// TIA Portal V20 export
// export: Created 2026-10-20T12:44:55.4293311Z, ExportSetting WithDefaults, DisplayName Totally Integrated Automation Portal, DisplayVersion V20 Update 6, DisplayName TIA Portal Openness, DisplayVersion V20 Update 6, DisplayName TIA Portal Version Control Interface, DisplayVersion V20 Update 6, DisplayName SINAMICS Startdrive Advanced, DisplayVersion V20 SP1, DisplayName SINAMICS Startdrive G130, G150, S120, S150, SINAMICS MV, G220, S200, S210, DisplayVersion V20 SP1, DisplayName SINAMICS Startdrive G110M, G120, G120C, G120D, G120P, G115D, DisplayVersion V20 SP1, DisplayName STEP 7 Professional, DisplayVersion V20 Update 6, DisplayName STEP 7 Safety, DisplayVersion V20 Update 2, DisplayName WinCC Basic/Comfort/Advanced, DisplayVersion V20 Update 6, DisplayName WinCC Unified, DisplayVersion V20 Update 6
FUNCTION "CNV_Selector_1" : Void   // FC60, SCL
{ S7_Optimized_Access := 'TRUE' }
VERSION : 0.1
// stored: AutoNumber true, IsIECCheckEnabled false, SetENOAutomatically false, UDAEnableTagReadback false
   VAR_INPUT
      Sys_No : UInt;
      Zone : UInt;
      CNV1_2_Selected : UInt;
   END_VAR
   VAR_OUTPUT
      ID : DInt;
      "ID(1)" : DInt;
   END_VAR
BEGIN
   //CNV SCREEN SELECTION
   CASE #Sys_No OF
       0:
           #ID := 0;
           #"ID(1)" := 0;

       1://SYSTEM 1
           #ID := "Settings_DB".ECnv_Sys[1].ID; // EXTRACTOR CONVEYOR
           CASE #Zone OF
               11: //LEVEL 1
                   IF #CNV1_2_Selected = 1 THEN
                       #"ID(1)" := "Settings_DB".LCnv_Sys[1].Cnv_Level[1].Cnv1.ID; //CNV 1
                   ELSIF #CNV1_2_Selected = 2 THEN
                       #"ID(1)" := "Settings_DB".LCnv_Sys[1].Cnv_Level[1].Cnv2.ID; //CNV 2
                   END_IF;
               12: //LEVEL 2
                   IF #CNV1_2_Selected = 1 THEN
                       #"ID(1)" := "Settings_DB".LCnv_Sys[1].Cnv_Level[2].Cnv1.ID; //CNV 1
                   ELSIF #CNV1_2_Selected = 2 THEN
                       #"ID(1)" := "Settings_DB".LCnv_Sys[1].Cnv_Level[2].Cnv2.ID; //CNV 2
                   END_IF;
               13: //LEVEL 3
                   IF #CNV1_2_Selected = 1 THEN
                       #"ID(1)" := "Settings_DB".LCnv_Sys[1].Cnv_Level[3].Cnv1.ID; //CNV 1
                   ELSIF #CNV1_2_Selected = 2 THEN
                       #"ID(1)" := "Settings_DB".LCnv_Sys[1].Cnv_Level[3].Cnv2.ID; //CNV 2
                   END_IF;
               14: //LEVEL 4
                   IF #CNV1_2_Selected = 1 THEN
                       #"ID(1)" := "Settings_DB".LCnv_Sys[1].Cnv_Level[4].Cnv1.ID; //CNV 1
                   ELSIF #CNV1_2_Selected = 2 THEN
                       #"ID(1)" := "Settings_DB".LCnv_Sys[1].Cnv_Level[4].Cnv2.ID; //CNV 2
                   END_IF;
               15: //LEVEL 5
                   IF #CNV1_2_Selected = 1 THEN
                       #"ID(1)" := "Settings_DB".LCnv_Sys[1].Cnv_Level[5].Cnv1.ID; //CNV 1
                   ELSIF #CNV1_2_Selected = 2 THEN
                       #"ID(1)" := "Settings_DB".LCnv_Sys[1].Cnv_Level[5].Cnv2.ID; //CNV 2
                   END_IF;
               16: //LEVEL 6
                   IF #CNV1_2_Selected = 1 THEN
                       #"ID(1)" := "Settings_DB".LCnv_Sys[1].Cnv_Level[6].Cnv1.ID; //CNV 1
                   ELSIF #CNV1_2_Selected = 2 THEN
                       #"ID(1)" := "Settings_DB".LCnv_Sys[1].Cnv_Level[6].Cnv2.ID; //CNV 2
                   END_IF;
               17: //LEVEL 7
                   IF #CNV1_2_Selected = 1 THEN
                       #"ID(1)" := "Settings_DB".LCnv_Sys[1].Cnv_Level[7].Cnv1.ID; //CNV 1
                   ELSIF #CNV1_2_Selected = 2 THEN
                       #"ID(1)" := "Settings_DB".LCnv_Sys[1].Cnv_Level[7].Cnv2.ID; //CNV 2
                   END_IF;
               18: //LEVEL 8
                   IF #CNV1_2_Selected = 1 THEN
                       #"ID(1)" := "Settings_DB".LCnv_Sys[1].Cnv_Level[8].Cnv1.ID; //CNV 1
                   ELSIF #CNV1_2_Selected = 2 THEN
                       #"ID(1)" := "Settings_DB".LCnv_Sys[1].Cnv_Level[8].Cnv2.ID; //CNV 2
                   END_IF;
               19: //LEVEL 1
                   IF #CNV1_2_Selected = 1 THEN
                       #"ID(1)" := "Settings_DB".LCnv_Sys[1].Cnv_Level[1].Cnv1.ID; //CNV 1
                   ELSIF #CNV1_2_Selected = 2 THEN
                       #"ID(1)" := "Settings_DB".LCnv_Sys[1].Cnv_Level[1].Cnv2.ID; //CNV 2
                   END_IF;
           END_CASE;

       2://SYSTEM 2
           #ID := "Settings_DB".ECnv_Sys[2].ID; // EXTRACTOR CONVEYOR
           CASE #Zone OF
               21: //LEVEL 1
                   IF #CNV1_2_Selected = 1 THEN
                       #"ID(1)" := "Settings_DB".LCnv_Sys[2].Cnv_Level[1].Cnv1.ID; //CNV 1
                   ELSIF #CNV1_2_Selected = 2 THEN
                       #"ID(1)" := "Settings_DB".LCnv_Sys[2].Cnv_Level[1].Cnv2.ID; //CNV 2
                   END_IF;
               22: //LEVEL 2
                   IF #CNV1_2_Selected = 1 THEN
                       #"ID(1)" := "Settings_DB".LCnv_Sys[2].Cnv_Level[2].Cnv1.ID; //CNV 1
                   ELSIF #CNV1_2_Selected = 2 THEN
                       #"ID(1)" := "Settings_DB".LCnv_Sys[2].Cnv_Level[2].Cnv2.ID; //CNV 2
                   END_IF;
               23: //LEVEL 3
                   IF #CNV1_2_Selected = 1 THEN
                       #"ID(1)" := "Settings_DB".LCnv_Sys[2].Cnv_Level[3].Cnv1.ID; //CNV 1
                   ELSIF #CNV1_2_Selected = 2 THEN
                       #"ID(1)" := "Settings_DB".LCnv_Sys[2].Cnv_Level[3].Cnv2.ID; //CNV 2
                   END_IF;
               24: //LEVEL 4
                   IF #CNV1_2_Selected = 1 THEN
                       #"ID(1)" := "Settings_DB".LCnv_Sys[2].Cnv_Level[4].Cnv1.ID; //CNV 1
                   ELSIF #CNV1_2_Selected = 2 THEN
                       #"ID(1)" := "Settings_DB".LCnv_Sys[2].Cnv_Level[4].Cnv2.ID; //CNV 2
                   END_IF;
               25: //LEVEL 5
                   IF #CNV1_2_Selected = 1 THEN
                       #"ID(1)" := "Settings_DB".LCnv_Sys[2].Cnv_Level[5].Cnv1.ID; //CNV 1
                   ELSIF #CNV1_2_Selected = 2 THEN
                       #"ID(1)" := "Settings_DB".LCnv_Sys[2].Cnv_Level[5].Cnv2.ID; //CNV 2
                   END_IF;
               26: //LEVEL 6
                   IF #CNV1_2_Selected = 1 THEN
                       #"ID(1)" := "Settings_DB".LCnv_Sys[2].Cnv_Level[6].Cnv1.ID; //CNV 1
                   ELSIF #CNV1_2_Selected = 2 THEN
                       #"ID(1)" := "Settings_DB".LCnv_Sys[2].Cnv_Level[6].Cnv2.ID; //CNV 2
                   END_IF;
               27: //LEVEL 7
                   IF #CNV1_2_Selected = 1 THEN
                       #"ID(1)" := "Settings_DB".LCnv_Sys[2].Cnv_Level[7].Cnv1.ID; //CNV 1
                   ELSIF #CNV1_2_Selected = 2 THEN
                       #"ID(1)" := "Settings_DB".LCnv_Sys[2].Cnv_Level[7].Cnv2.ID; //CNV 2
                   END_IF;
               28: //LEVEL 8
                   IF #CNV1_2_Selected = 1 THEN
                       #"ID(1)" := "Settings_DB".LCnv_Sys[2].Cnv_Level[8].Cnv1.ID; //CNV 1
                   ELSIF #CNV1_2_Selected = 2 THEN
                       #"ID(1)" := "Settings_DB".LCnv_Sys[2].Cnv_Level[8].Cnv2.ID; //CNV 2
                   END_IF;
               29: //LEVEL 1
                   IF #CNV1_2_Selected = 1 THEN
                       #"ID(1)" := "Settings_DB".LCnv_Sys[2].Cnv_Level[1].Cnv1.ID; //CNV 1
                   ELSIF #CNV1_2_Selected = 2 THEN
                       #"ID(1)" := "Settings_DB".LCnv_Sys[2].Cnv_Level[1].Cnv2.ID; //CNV 2
                   END_IF;
           END_CASE;

       3://SYSTEM 3
           #ID := "Settings_DB".ECnv_Sys[3].ID; // EXTRACTOR CONVEYOR
           CASE #Zone OF
               31: //LEVEL 1
                   IF #CNV1_2_Selected = 1 THEN
                       #"ID(1)" := "Settings_DB".LCnv_Sys[3].Cnv_Level[1].Cnv1.ID; //CNV 1
                   ELSIF #CNV1_2_Selected = 2 THEN
                       #"ID(1)" := "Settings_DB".LCnv_Sys[3].Cnv_Level[1].Cnv2.ID; //CNV 2
                   END_IF;
               32: //LEVEL 2
                   IF #CNV1_2_Selected = 1 THEN
                       #"ID(1)" := "Settings_DB".LCnv_Sys[3].Cnv_Level[2].Cnv1.ID; //CNV 1
                   ELSIF #CNV1_2_Selected = 2 THEN
                       #"ID(1)" := "Settings_DB".LCnv_Sys[3].Cnv_Level[2].Cnv2.ID; //CNV 2
                   END_IF;
               33: //LEVEL 3
                   IF #CNV1_2_Selected = 1 THEN
                       #"ID(1)" := "Settings_DB".LCnv_Sys[3].Cnv_Level[3].Cnv1.ID; //CNV 1
                   ELSIF #CNV1_2_Selected = 2 THEN
                       #"ID(1)" := "Settings_DB".LCnv_Sys[3].Cnv_Level[3].Cnv2.ID; //CNV 2
                   END_IF;
               34: //LEVEL 4
                   IF #CNV1_2_Selected = 1 THEN
                       #"ID(1)" := "Settings_DB".LCnv_Sys[3].Cnv_Level[4].Cnv1.ID; //CNV 1
                   ELSIF #CNV1_2_Selected = 2 THEN
                       #"ID(1)" := "Settings_DB".LCnv_Sys[3].Cnv_Level[4].Cnv2.ID; //CNV 2
                   END_IF;
               35: //LEVEL 5
                   IF #CNV1_2_Selected = 1 THEN
                       #"ID(1)" := "Settings_DB".LCnv_Sys[3].Cnv_Level[5].Cnv1.ID; //CNV 1
                   ELSIF #CNV1_2_Selected = 2 THEN
                       #"ID(1)" := "Settings_DB".LCnv_Sys[3].Cnv_Level[5].Cnv2.ID; //CNV 2
                   END_IF;
               36: //LEVEL 6
                   IF #CNV1_2_Selected = 1 THEN
                       #"ID(1)" := "Settings_DB".LCnv_Sys[3].Cnv_Level[6].Cnv1.ID; //CNV 1
                   ELSIF #CNV1_2_Selected = 2 THEN
                       #"ID(1)" := "Settings_DB".LCnv_Sys[3].Cnv_Level[6].Cnv2.ID; //CNV 2
                   END_IF;
               37: //LEVEL 7
                   IF #CNV1_2_Selected = 1 THEN
                       #"ID(1)" := "Settings_DB".LCnv_Sys[3].Cnv_Level[7].Cnv1.ID; //CNV 1
                   ELSIF #CNV1_2_Selected = 2 THEN
                       #"ID(1)" := "Settings_DB".LCnv_Sys[3].Cnv_Level[7].Cnv2.ID; //CNV 2
                   END_IF;
               38: //LEVEL 8
                   IF #CNV1_2_Selected = 1 THEN
                       #"ID(1)" := "Settings_DB".LCnv_Sys[3].Cnv_Level[8].Cnv1.ID; //CNV 1
                   ELSIF #CNV1_2_Selected = 2 THEN
                       #"ID(1)" := "Settings_DB".LCnv_Sys[3].Cnv_Level[8].Cnv2.ID; //CNV 2
                   END_IF;
               39: //LEVEL 1
                   IF #CNV1_2_Selected = 1 THEN
                       #"ID(1)" := "Settings_DB".LCnv_Sys[3].Cnv_Level[1].Cnv1.ID; //CNV 1
                   ELSIF #CNV1_2_Selected = 2 THEN
                       #"ID(1)" := "Settings_DB".LCnv_Sys[3].Cnv_Level[1].Cnv2.ID; //CNV 2
                   END_IF;
           END_CASE;

       4://SYSTEM 4
           #ID := "Settings_DB".ECnv_Sys[4].ID; // EXTRACTOR CONVEYOR
           CASE #Zone OF
               41: //LEVEL 1
                   IF #CNV1_2_Selected = 1 THEN
                       #"ID(1)" := "Settings_DB".LCnv_Sys[4].Cnv_Level[1].Cnv1.ID; //CNV 1
                   ELSIF #CNV1_2_Selected = 2 THEN
                       #"ID(1)" := "Settings_DB".LCnv_Sys[4].Cnv_Level[1].Cnv2.ID; //CNV 2
                   END_IF;
               42: //LEVEL 2
                   IF #CNV1_2_Selected = 1 THEN
                       #"ID(1)" := "Settings_DB".LCnv_Sys[4].Cnv_Level[2].Cnv1.ID; //CNV 1
                   ELSIF #CNV1_2_Selected = 2 THEN
                       #"ID(1)" := "Settings_DB".LCnv_Sys[4].Cnv_Level[2].Cnv2.ID; //CNV 2
                   END_IF;
               43: //LEVEL 3
                   IF #CNV1_2_Selected = 1 THEN
                       #"ID(1)" := "Settings_DB".LCnv_Sys[4].Cnv_Level[3].Cnv1.ID; //CNV 1
                   ELSIF #CNV1_2_Selected = 2 THEN
                       #"ID(1)" := "Settings_DB".LCnv_Sys[4].Cnv_Level[3].Cnv2.ID; //CNV 2
                   END_IF;
               44: //LEVEL 4
                   IF #CNV1_2_Selected = 1 THEN
                       #"ID(1)" := "Settings_DB".LCnv_Sys[4].Cnv_Level[4].Cnv1.ID; //CNV 1
                   ELSIF #CNV1_2_Selected = 2 THEN
                       #"ID(1)" := "Settings_DB".LCnv_Sys[4].Cnv_Level[4].Cnv2.ID; //CNV 2
                   END_IF;
               45: //LEVEL 5
                   IF #CNV1_2_Selected = 1 THEN
                       #"ID(1)" := "Settings_DB".LCnv_Sys[4].Cnv_Level[5].Cnv1.ID; //CNV 1
                   ELSIF #CNV1_2_Selected = 2 THEN
                       #"ID(1)" := "Settings_DB".LCnv_Sys[4].Cnv_Level[5].Cnv2.ID; //CNV 2
                   END_IF;
               46: //LEVEL 6
                   IF #CNV1_2_Selected = 1 THEN
                       #"ID(1)" := "Settings_DB".LCnv_Sys[4].Cnv_Level[6].Cnv1.ID; //CNV 1
                   ELSIF #CNV1_2_Selected = 2 THEN
                       #"ID(1)" := "Settings_DB".LCnv_Sys[4].Cnv_Level[6].Cnv2.ID; //CNV 2
                   END_IF;
               47: //LEVEL 7
                   IF #CNV1_2_Selected = 1 THEN
                       #"ID(1)" := "Settings_DB".LCnv_Sys[4].Cnv_Level[7].Cnv1.ID; //CNV 1
                   ELSIF #CNV1_2_Selected = 2 THEN
                       #"ID(1)" := "Settings_DB".LCnv_Sys[4].Cnv_Level[7].Cnv2.ID; //CNV 2
                   END_IF;
               48: //LEVEL 8
                   IF #CNV1_2_Selected = 1 THEN
                       #"ID(1)" := "Settings_DB".LCnv_Sys[4].Cnv_Level[8].Cnv1.ID; //CNV 1
                   ELSIF #CNV1_2_Selected = 2 THEN
                       #"ID(1)" := "Settings_DB".LCnv_Sys[4].Cnv_Level[8].Cnv2.ID; //CNV 2
                   END_IF;
               49: //LEVEL 1
                   IF #CNV1_2_Selected = 1 THEN
                       #"ID(1)" := "Settings_DB".LCnv_Sys[4].Cnv_Level[1].Cnv1.ID; //CNV 1
                   ELSIF #CNV1_2_Selected = 2 THEN
                       #"ID(1)" := "Settings_DB".LCnv_Sys[4].Cnv_Level[1].Cnv2.ID; //CNV 2
                   END_IF;
           END_CASE;

       5://SYSTEM 5
           #ID := "Settings_DB".ECnv_Sys[5].ID; // EXTRACTOR CONVEYOR
           CASE #Zone OF
               51: //LEVEL 1
                   IF #CNV1_2_Selected = 1 THEN
                       #"ID(1)" := "Settings_DB".LCnv_Sys[5].Cnv_Level[1].Cnv1.ID; //CNV 1
                   ELSIF #CNV1_2_Selected = 2 THEN
                       #"ID(1)" := "Settings_DB".LCnv_Sys[5].Cnv_Level[1].Cnv2.ID; //CNV 2
                   END_IF;
               52: //LEVEL 2
                   IF #CNV1_2_Selected = 1 THEN
                       #"ID(1)" := "Settings_DB".LCnv_Sys[5].Cnv_Level[2].Cnv1.ID; //CNV 1
                   ELSIF #CNV1_2_Selected = 2 THEN
                       #"ID(1)" := "Settings_DB".LCnv_Sys[5].Cnv_Level[2].Cnv2.ID; //CNV 2
                   END_IF;
               53: //LEVEL 3
                   IF #CNV1_2_Selected = 1 THEN
                       #"ID(1)" := "Settings_DB".LCnv_Sys[5].Cnv_Level[3].Cnv1.ID; //CNV 1
                   ELSIF #CNV1_2_Selected = 2 THEN
                       #"ID(1)" := "Settings_DB".LCnv_Sys[5].Cnv_Level[3].Cnv2.ID; //CNV 2
                   END_IF;
               54: //LEVEL 4
                   IF #CNV1_2_Selected = 1 THEN
                       #"ID(1)" := "Settings_DB".LCnv_Sys[5].Cnv_Level[4].Cnv1.ID; //CNV 1
                   ELSIF #CNV1_2_Selected = 2 THEN
                       #"ID(1)" := "Settings_DB".LCnv_Sys[5].Cnv_Level[4].Cnv2.ID; //CNV 2
                   END_IF;
               55: //LEVEL 5
                   IF #CNV1_2_Selected = 1 THEN
                       #"ID(1)" := "Settings_DB".LCnv_Sys[5].Cnv_Level[5].Cnv1.ID; //CNV 1
                   ELSIF #CNV1_2_Selected = 2 THEN
                       #"ID(1)" := "Settings_DB".LCnv_Sys[5].Cnv_Level[5].Cnv2.ID; //CNV 2
                   END_IF;
               56: //LEVEL 6
                   IF #CNV1_2_Selected = 1 THEN
                       #"ID(1)" := "Settings_DB".LCnv_Sys[5].Cnv_Level[6].Cnv1.ID; //CNV 1
                   ELSIF #CNV1_2_Selected = 2 THEN
                       #"ID(1)" := "Settings_DB".LCnv_Sys[5].Cnv_Level[6].Cnv2.ID; //CNV 2
                   END_IF;
               57: //LEVEL 7
                   IF #CNV1_2_Selected = 1 THEN
                       #"ID(1)" := "Settings_DB".LCnv_Sys[5].Cnv_Level[7].Cnv1.ID; //CNV 1
                   ELSIF #CNV1_2_Selected = 2 THEN
                       #"ID(1)" := "Settings_DB".LCnv_Sys[5].Cnv_Level[7].Cnv2.ID; //CNV 2
                   END_IF;
               58: //LEVEL 8
                   IF #CNV1_2_Selected = 1 THEN
                       #"ID(1)" := "Settings_DB".LCnv_Sys[5].Cnv_Level[8].Cnv1.ID; //CNV 1
                   ELSIF #CNV1_2_Selected = 2 THEN
                       #"ID(1)" := "Settings_DB".LCnv_Sys[5].Cnv_Level[8].Cnv2.ID; //CNV 2
                   END_IF;
               59: //LEVEL 1
                   IF #CNV1_2_Selected = 1 THEN
                       #"ID(1)" := "Settings_DB".LCnv_Sys[5].Cnv_Level[1].Cnv1.ID; //CNV 1
                   ELSIF #CNV1_2_Selected = 2 THEN
                       #"ID(1)" := "Settings_DB".LCnv_Sys[5].Cnv_Level[1].Cnv2.ID; //CNV 2
                   END_IF;
           END_CASE;
   END_CASE;
END_FUNCTION
